FUNCTION_BLOCK FB_ProdRecipe_Manage
VAR_INPUT
END_VAR
VAR_OUTPUT
END_VAR
VAR
	stProdParam_HMI: ST_Production_Parameter;

	bReInit: BOOL;
END_VAR

IF bReInit THEN;
	FB_INIT(bInCopyCode:=FALSE,bInitRetains:=FALSE);
	bReInit:=FALSE;
	//FB_INIT.bInitRetains:=TRUE;
END_IF
mPercentage_Calculation();
mGet_Recipe_list();

g_Prod.dtProdTimeMin:=dtRealTime-T#2H;
g_Prod.dtProdTimeMax:=dtRealTime+T#7D;

METHOD FB_INIT : BOOL
VAR_INPUT
END_VAR
VAR_INPUT
    bInitRetains : BOOL; // TRUE if the FB is being initialized after a warm restart
    bInCopyCode : BOOL;  // TRUE if the FB is being initialized in copy code
END_VAR
VAR
	i: INT;
	k: INT;
END_VAR
FOR i:=0 TO g_Prod.cMax_Prod_Recipe DO
	
	g_Prod.arrRecipeMarinade[i].prodType:=E_Prod_Type.Marinade;
	g_Prod.arrRecipeColor[i].prodType:=E_Prod_Type.Color;
	
	g_Prod.arrRecipeMarinade[i].arr_Component[1].sDescription:='Water';
	g_Prod.arrRecipeColor[i].arr_Component[1].sDescription:='Water';
	
	g_Prod.arrRecipeMarinade[i].arr_Component[1].eIngredientType:=E_Ingredient_type.eWater;
	g_Prod.arrRecipeColor[i].arr_Component[1].eIngredientType:=E_Ingredient_type.eWater;

	FOR k:=2 TO g_Prod.cMaxCompInProduct-1 DO
		//g_Prod.arrRecipeMarinade[i].arr_Component[k].sDescription:='Powder';
		//g_Prod.arrRecipeColor[i].arr_Component[k].sDescription:='Powder';
		
		g_Prod.arrRecipeMarinade[i].arr_Component[k].eIngredientType:=E_Ingredient_type.ePowder;
		g_Prod.arrRecipeColor[i].arr_Component[k].eIngredientType:=E_Ingredient_type.ePowder;		
	END_FOR
	
	
	
	g_Prod.arrRecipeMarinade[i].arr_Component[10].sDescription:='Oil';
	g_Prod.arrRecipeColor[i].arr_Component[10].sDescription:='Oil';
	
	g_Prod.arrRecipeMarinade[i].arr_Component[10].eIngredientType:=E_Ingredient_type.eOil;
	g_Prod.arrRecipeColor[i].arr_Component[10].eIngredientType:=E_Ingredient_type.eOil;	

END_FOR
END_METHOD

METHOD mGet_Recipe_list : BOOL
VAR_INPUT
END_VAR

VAR
	i: INT;
END_VAR
FOR i:=1 TO g_Prod.cMax_Prod_Recipe DO
	g_Prod.listRecipe_Marinade[i]:=g_Prod.arrRecipeMarinade[i].Description;
	g_Prod.listRecipe_Color[i]:=g_Prod.arrRecipeColor[i].Description;
	
	
END_FOR
END_METHOD

METHOD mPercentage_Calculation : BOOL
VAR_INPUT
END_VAR

VAR
	i: INT;
	tempPercentage_M: REAL;
	tempPercentage_C: REAL;
	k: INT;
END_VAR

FOR i:=1 TO g_Prod.cMax_Prod_Recipe DO
	tempPercentage_M:=0;
	tempPercentage_C:=0;	
	FOR k:=2 TO g_Prod.cMaxCompInProduct DO
		tempPercentage_M:=tempPercentage_M + g_Prod.arrRecipeMarinade[i].arr_Component[k].rWeightPercentage;
		tempPercentage_C:=tempPercentage_C + g_Prod.arrRecipeColor[i].arr_Component[k].rWeightPercentage;
	END_FOR
	g_Prod.arrRecipeMarinade[i].arr_Component[1].rWeightPercentage:=100-tempPercentage_M;
	g_Prod.arrRecipeColor[i].arr_Component[1].rWeightPercentage:=100-tempPercentage_C;
END_FOR
END_METHOD

END_FUNCTION_BLOCK

(* stored: Version 1.1.0.1, ProductVersion 3.1.4024.15
   POU FB_ProdRecipe_Manage: Id {6d224ab8-fc12-45df-bf04-9b71c4fddbfa}, SpecialFunc None
   Method FB_INIT: Id {829a4d5a-b2e2-488a-be22-05f2cbbb07cb}
   Method mGet_Recipe_list: Id {86031595-6db8-40d6-a74f-31cac555018a}
   Method mPercentage_Calculation: Id {f4c275b1-d3ea-444b-987c-802362ed0562} *)
